(*
SPDX-FileCopyrightText: © 2026 Oleksandr Tiutyk <trofimich@gmail.com>
SPDX-License-Identifier: MIT
License: https://opensource.org/license/mit
*)

(*!
<summary>Separates filesystem scenario execution from cleanup and result reporting.</summary>
<description>
A case remains active while cleanup is pending. Completed drain and cleanup attempts permit FINISHED
and result reporting. Errors remain test failures and do not authorize deleting unowned paths.
Cleanup has no forced deadline. These phases do not guarantee physical close after a native release failure.
</description>
*)
{attribute 'qualified_only'}
{attribute 'strict'}
TYPE FILE_TEST_LIFECYCLE :
(
	//! <summary>Advance the scenario and its deadline until its normal or failed outcome is known.</summary>
	RUNNING_SCENARIO,
	//! <summary>Keep the case active while retained resources stop and owned cleanup attempts finish.</summary>
	CLEANING_UP,
	//! <summary>Cleanup observations were reported for this run.</summary>
	FINISHED
);
END_TYPE

(* stored: Version 1.1.0.1
   DUT FILE_TEST_LIFECYCLE: Id {fe324de8-d781-4a3e-a68b-2b1fad78b77a} *)
